// POUs/_FB_ConfigMachine
(****************************************************************************************************<br>
© Syntegon Group.<br>
All rights reserved, also regarding any disposal, exploitation, reproduction, editing, distribution,<br>
as well as in the event of applications for industrial property rights.<br>
*****************************************************************************************************<br>
DESCRIPTION:<br>
The machine as a whole (config protocol 3, ADR 0022): the recipe fields the application declares (process values<br>
such as belt speed, picks per cycle, the product pattern), their staging by the Simulator with the mechanism of the<br>
parameter sets, and the machine commands Start, Stop and Reset the application answers. One per application,<br>
listed in the config manifest with id 0. Typical cycle:<br>
  fb_Machine.m_Register(vio_Manifest := GVL_Config.stManifest, vi_udn_Id := 0);<br>
  fb_Machine.m_DeclareField(vi_un_Field := 1, vi_str_Name := 'BeltSpeed', vi_udn_Group := fb_Infeed.m_Id(),<br>
    vi_e_Type := E_ConfigFieldType.NUMBER, vi_str_Unit := 'mm/s', vi_lr_Min := 0, vi_lr_Max := 500,<br>
    vi_lr_ProgramValue := 150);<br>
  fb_Machine.m_SetText(vi_un_Field := 1, vi_str_Label := 'Belt speed', vi_str_Description := 'Speed of the infeed');<br>
  fb_Machine.m_SetVisibleWhen(vi_un_Field := 3, vi_un_OnField := 2, vi_dn_Value := 0);  // field 3 only with 2 = 0<br>
  fb_Machine.m_Cycle(vio_Set := RecipeSet, vi_b_ApplyAllowed := b_Stopped);<br>
  lr_BeltSpeed := fb_Machine.m_Value(vi_un_Field := 1);<br>
  CASE fb_Machine.m_Command() OF E_ConfigCommand.START: ...<br>
    fb_Machine.m_AnswerCommand(vi_b_Accepted := TRUE, vi_str_Reason := ''); END_CASE<br>
RecipeSet is the application's VAR PERSISTENT ST_ConfigRecipeSet.<br>
*****************************************************************************************************<br>
OUTPUT VALUES:<br>
vo_Config is the contract structure the gateway reads and writes at the path in the config manifest.<br>
*****************************************************************************************************<br>
LIMITS:<br>
CONFIG_un_MAX_RECIPE_FIELDS fields, CONFIG_un_MAX_CHOICES choices each. The gateway reads the declarations when<br>
it discovers the PLC: declare every field from the start and keep their order.<br>
*****************************************************************************************************<br>
VERSION         ¦ DATE       ¦ NAME      ¦ CHANGE<br>
Syn_Config 2.1.0 ¦ 2026-11-14 ¦ J.Willner ¦ Created: recipe fields and machine commands (protocol 3)<br>
Syn_Config 2.2.0 ¦ 2026-11-14 ¦ J.Willner ¦ m_SetText, m_SetVisibleWhen (protocol 4, #49)<br>
Syn_Config 2.3.0 ¦ 2026-11-14 ¦ J.Willner ¦ m_Cycle through m_HandleStaging<br>
****************************************************************************************************)
FUNCTION_BLOCK _FB_ConfigMachine EXTENDS _FB_ConfigComponent
VAR_OUTPUT
	vo_Config							: ST_ConfigMachine;	// contract structure of the gateway
END_VAR

(****************************************************************************************************<br>
© Syntegon Group.<br>
All rights reserved, also regarding any disposal, exploitation, reproduction, editing, distribution,<br>
as well as in the event of applications for industrial property rights.<br>
*****************************************************************************************************<br>
DESCRIPTION:<br>
Answers the waiting machine command: accepted, or rejected with the reason the Simulator shows. The command no<br>
longer waits afterwards.<br>
*****************************************************************************************************<br>
OUTPUT VALUES:<br>
FALSE while no command waits.<br>
****************************************************************************************************)
METHOD m_AnswerCommand : BOOL
VAR_INPUT
	vi_b_Accepted						: BOOL;	// TRUE: the application carries the command out
	vi_str_Reason						: STRING(80);	// why it is rejected, '' when accepted
END_VAR
m_AnswerCommand := vo_Config.stCommand.bRequested;
IF NOT m_AnswerCommand THEN
	RETURN;
END_IF
vo_Config.stCommandStatus.nHandledCommandId := vo_Config.stCommand.nCommandId;
vo_Config.stCommandStatus.eResult := SEL(vi_b_Accepted, E_ConfigCommandResult.REJECTED, E_ConfigCommandResult.ACCEPTED);
vo_Config.stCommandStatus.sMessage := SEL(vi_b_Accepted, vi_str_Reason, '');
vo_Config.stCommand.bRequested := FALSE;
END_METHOD

(****************************************************************************************************<br>
© Syntegon Group.<br>
All rights reserved, also regarding any disposal, exploitation, reproduction, editing, distribution,<br>
as well as in the event of applications for industrial property rights.<br>
*****************************************************************************************************<br>
DESCRIPTION:<br>
The machine command waiting for the application's answer (START, STOP, RESET); NONE while none waits. Answer it<br>
with m_AnswerCommand: the application alone decides whether it is carried out.<br>
****************************************************************************************************)
METHOD m_Command : E_ConfigCommand
IF vo_Config.stCommand.bRequested THEN
	m_Command := vo_Config.stCommand.eCommand;
ELSE
	m_Command := E_ConfigCommand.NONE;
END_IF
END_METHOD

(****************************************************************************************************<br>
© Syntegon Group.<br>
All rights reserved, also regarding any disposal, exploitation, reproduction, editing, distribution,<br>
as well as in the event of applications for industrial property rights.<br>
*****************************************************************************************************<br>
DESCRIPTION:<br>
Every cycle, after the fields are declared: handles a staged recipe or a reset (a recipe only while<br>
vi_b_ApplyAllowed), keeps the active recipe in vio_Set and gives the effective values in vo_Config.aActive: the<br>
active recipe while one is valid, else the fields' program values.<br>
*****************************************************************************************************<br>
OUTPUT VALUES:<br>
TRUE in the cycle a recipe was taken over or reset.<br>
****************************************************************************************************)
METHOD m_Cycle : BOOL
VAR_IN_OUT
	vio_Set								: ST_ConfigRecipeSet;	// the application's VAR PERSISTENT active recipe
END_VAR
VAR_INPUT
	vi_b_ApplyAllowed					: BOOL;	// [-] a staged recipe may be taken over now, e.g. while the machine stands
END_VAR
VAR
	b_TempTakeOver						: BOOL;	// the staged recipe was taken over: copy it
	un_TempIndex						: UINT;
END_VAR
m_Cycle := m_HandleStaging(vio_Staging := vo_Config.stStaging, vio_Status := vo_Config.stStatus, vio_b_Valid := vio_Set.bValid,
	vio_udn_Version := vio_Set.nVersion, vio_udn_LastVersion := vio_Set.nLastVersion, vi_b_ApplyAllowed := vi_b_ApplyAllowed,
	vo_b_TakeOver => b_TempTakeOver);
IF b_TempTakeOver THEN
	vio_Set.aValues := vo_Config.aStaged;
END_IF


(****************************************************************************************************
EFFECTIVE VALUES
****************************************************************************************************)
un_TempIndex := 0;
WHILE un_TempIndex < vo_Config.nFieldCount AND un_TempIndex < CONFIG_GlobalConst_Param.CONFIG_un_MAX_RECIPE_FIELDS DO
	vo_Config.aActive[un_TempIndex] := SEL(vio_Set.bValid, vo_Config.aFields[un_TempIndex].fProgramValue,
		vio_Set.aValues[un_TempIndex]);
	un_TempIndex := un_TempIndex + 1;
END_WHILE
END_METHOD

(****************************************************************************************************<br>
© Syntegon Group.<br>
All rights reserved, also regarding any disposal, exploitation, reproduction, editing, distribution,<br>
as well as in the event of applications for industrial property rights.<br>
*****************************************************************************************************<br>
DESCRIPTION:<br>
Declares recipe field vi_un_Field (1..CONFIG_un_MAX_RECIPE_FIELDS): its name, the component it belongs to, how its<br>
value is kept, its unit, range and the program value that applies while no recipe is active. Fields are listed up<br>
to the highest one declared. Idempotent: call it every cycle, before m_Cycle. A CHOICE field's values are named with<br>
m_SetChoice and range from 0; its vi_lr_Min and vi_lr_Max are not used, nor a SWITCH's.<br>
*****************************************************************************************************<br>
OUTPUT VALUES:<br>
FALSE for vi_un_Field = 0 or above CONFIG_un_MAX_RECIPE_FIELDS.<br>
****************************************************************************************************)
METHOD m_DeclareField : BOOL
VAR_INPUT
	vi_un_Field							: UINT;	// [-] 1..CONFIG_un_MAX_RECIPE_FIELDS
	vi_str_Name							: STRING(31);	// unique in the recipe, e.g. 'BeltSpeed'
	vi_udn_Group						: UDINT;	// [-] manifest id of the Syn_Visu component, 0 = the whole machine
	vi_e_Type							: E_ConfigFieldType;
	vi_str_Unit							: STRING(15);	// e.g. 'mm/s', '' = none
	vi_lr_Min							: LREAL;	// smallest value of a NUMBER or INTEGER field
	vi_lr_Max							: LREAL;	// largest value of a NUMBER or INTEGER field
	vi_lr_ProgramValue					: LREAL;	// the application's own value; a SWITCH: 1 = on
END_VAR
m_DeclareField := vi_un_Field > 0 AND vi_un_Field <= CONFIG_GlobalConst_Param.CONFIG_un_MAX_RECIPE_FIELDS;
IF NOT m_DeclareField THEN
	RETURN;
END_IF
vo_Config.aFields[vi_un_Field - 1].sName := vi_str_Name;
vo_Config.aFields[vi_un_Field - 1].nGroup := vi_udn_Group;
vo_Config.aFields[vi_un_Field - 1].eType := vi_e_Type;
vo_Config.aFields[vi_un_Field - 1].sUnit := vi_str_Unit;
vo_Config.aFields[vi_un_Field - 1].fMin := vi_lr_Min;
vo_Config.aFields[vi_un_Field - 1].fMax := vi_lr_Max;
vo_Config.aFields[vi_un_Field - 1].fProgramValue := vi_lr_ProgramValue;
IF vi_un_Field > vo_Config.nFieldCount THEN
	vo_Config.nFieldCount := vi_un_Field;
END_IF
END_METHOD

(****************************************************************************************************<br>
© Syntegon Group.<br>
All rights reserved, also regarding any disposal, exploitation, reproduction, editing, distribution,<br>
as well as in the event of applications for industrial property rights.<br>
*****************************************************************************************************<br>
DESCRIPTION:<br>
Effective value of an INTEGER or CHOICE recipe field as a whole number (see m_Value).<br>
****************************************************************************************************)
METHOD m_Integer : DINT
VAR_INPUT
	vi_un_Field							: UINT;	// [-] 1..the field count
END_VAR
m_Integer := LREAL_TO_DINT(m_Value(vi_un_Field := vi_un_Field));
END_METHOD

(****************************************************************************************************<br>
© Syntegon Group.<br>
All rights reserved, also regarding any disposal, exploitation, reproduction, editing, distribution,<br>
as well as in the event of applications for industrial property rights.<br>
*****************************************************************************************************<br>
DESCRIPTION:<br>
Why the staged recipe cannot be taken over; '' when it can: a value outside its field's range (NUMBER, INTEGER),<br>
not one of its choices (CHOICE), not a whole number (INTEGER, CHOICE) or not 0 or 1 (SWITCH).<br>
****************************************************************************************************)
METHOD PROTECTED m_InvalidStaged : STRING(80)
VAR
	un_TempIndex						: UINT;
	lr_TempValue						: LREAL;
	lr_TempMin							: LREAL;
	lr_TempMax							: LREAL;
END_VAR
m_InvalidStaged := '';
un_TempIndex := 0;
WHILE un_TempIndex < vo_Config.nFieldCount AND un_TempIndex < CONFIG_GlobalConst_Param.CONFIG_un_MAX_RECIPE_FIELDS DO
	lr_TempValue := vo_Config.aStaged[un_TempIndex];
	CASE vo_Config.aFields[un_TempIndex].eType OF
		E_ConfigFieldType.SWITCH:
			lr_TempMin := 0;
			lr_TempMax := 1;
		E_ConfigFieldType.CHOICE:
			lr_TempMin := 0;
			lr_TempMax := UINT_TO_LREAL(vo_Config.aFields[un_TempIndex].nChoiceCount) - 1;
	ELSE
		lr_TempMin := vo_Config.aFields[un_TempIndex].fMin;
		lr_TempMax := vo_Config.aFields[un_TempIndex].fMax;
	END_CASE
	(* The range first: only a value in range is turned into a whole number. NaN equals nothing, not even itself. *)
	IF lr_TempValue <> lr_TempValue OR lr_TempValue < lr_TempMin OR lr_TempValue > lr_TempMax THEN
		m_InvalidStaged := CONCAT(CONCAT('Field ', vo_Config.aFields[un_TempIndex].sName), CONCAT(': ', CONCAT(LREAL_TO_STRING(lr_TempValue),
			CONCAT(' is outside ', CONCAT(LREAL_TO_STRING(lr_TempMin), CONCAT(' to ', LREAL_TO_STRING(lr_TempMax)))))));
		RETURN;
	END_IF
	IF vo_Config.aFields[un_TempIndex].eType <> E_ConfigFieldType.NUMBER
		AND LINT_TO_LREAL(LREAL_TO_LINT(lr_TempValue)) <> lr_TempValue
	THEN
		m_InvalidStaged := CONCAT(CONCAT('Field ', vo_Config.aFields[un_TempIndex].sName), CONCAT(': ',
			CONCAT(LREAL_TO_STRING(lr_TempValue), ' is not a value of its type')));
		RETURN;
	END_IF
	un_TempIndex := un_TempIndex + 1;
END_WHILE
END_METHOD

(****************************************************************************************************<br>
© Syntegon Group.<br>
All rights reserved, also regarding any disposal, exploitation, reproduction, editing, distribution,<br>
as well as in the event of applications for industrial property rights.<br>
*****************************************************************************************************<br>
DESCRIPTION:<br>
Names value vi_un_Value (0..CONFIG_un_MAX_CHOICES-1) of the CHOICE field vi_un_Field, e.g. 0 = 'Lanes'. The field<br>
has as many choices as the highest value named plus one. Idempotent: call it every cycle with m_DeclareField.<br>
*****************************************************************************************************<br>
OUTPUT VALUES:<br>
FALSE for a field not declared or a value above CONFIG_un_MAX_CHOICES - 1.<br>
****************************************************************************************************)
METHOD m_SetChoice : BOOL
VAR_INPUT
	vi_un_Field							: UINT;	// [-] the field, 1..its count
	vi_un_Value							: UINT;	// [-] the value it names, from 0
	vi_str_Text							: STRING(31);	// e.g. 'Lanes'
END_VAR
m_SetChoice := vi_un_Field > 0 AND vi_un_Field <= vo_Config.nFieldCount
	AND vi_un_Value < CONFIG_GlobalConst_Param.CONFIG_un_MAX_CHOICES;
IF NOT m_SetChoice THEN
	RETURN;
END_IF
vo_Config.aFields[vi_un_Field - 1].aChoices[vi_un_Value] := vi_str_Text;
IF vi_un_Value >= vo_Config.aFields[vi_un_Field - 1].nChoiceCount THEN
	vo_Config.aFields[vi_un_Field - 1].nChoiceCount := vi_un_Value + 1;
END_IF
END_METHOD

(****************************************************************************************************<br>
© Syntegon Group.<br>
All rights reserved, also regarding any disposal, exploitation, reproduction, editing, distribution,<br>
as well as in the event of applications for industrial property rights.<br>
*****************************************************************************************************<br>
DESCRIPTION:<br>
Gives the declared field vi_un_Field the label the Simulator shows instead of its name put into words, and a<br>
description of what it is for, shown in the field's tooltip (config protocol 4, #49). Free text in the operators'<br>
language; the name stays the field's key. Idempotent: call it every cycle with m_DeclareField.<br>
*****************************************************************************************************<br>
OUTPUT VALUES:<br>
FALSE for a field not declared.<br>
****************************************************************************************************)
METHOD m_SetText : BOOL
VAR_INPUT
	vi_un_Field							: UINT;	// [-] the field, 1..its count
	vi_str_Label						: STRING(40);	// e.g. 'Belt speed', '' = the name put into words
	vi_str_Description					: STRING(160);	// what the field is for, '' = none
END_VAR
m_SetText := vi_un_Field > 0 AND vi_un_Field <= vo_Config.nFieldCount;
IF NOT m_SetText THEN
	RETURN;
END_IF
vo_Config.aFields[vi_un_Field - 1].sLabel := vi_str_Label;
vo_Config.aFields[vi_un_Field - 1].sDescription := vi_str_Description;
END_METHOD

(****************************************************************************************************<br>
© Syntegon Group.<br>
All rights reserved, also regarding any disposal, exploitation, reproduction, editing, distribution,<br>
as well as in the event of applications for industrial property rights.<br>
*****************************************************************************************************<br>
DESCRIPTION:<br>
Shows the declared field vi_un_Field in the Simulator only while field vi_un_OnField has the value vi_dn_Value<br>
(config protocol 4, #49), e.g. a lane count only while the pattern is Lanes. vi_un_OnField must be a SWITCH (0 / 1),<br>
CHOICE or INTEGER field and may belong to another group; a field depending on a hidden one is hidden too. A hidden<br>
field keeps its value and is written with the recipe. vi_un_OnField = 0 shows the field always. The gateway reports<br>
a condition on a NUMBER field, on the field itself, on a field not declared, on a value that field can never have<br>
or in a ring as a discovery error and shows that field always. Idempotent: call it every cycle with m_DeclareField.<br>
*****************************************************************************************************<br>
OUTPUT VALUES:<br>
FALSE for a field not declared.<br>
****************************************************************************************************)
METHOD m_SetVisibleWhen : BOOL
VAR_INPUT
	vi_un_Field							: UINT;	// [-] the field shown on condition, 1..its count
	vi_un_OnField						: UINT;	// [-] the field the condition reads, 0 = always shown
	vi_dn_Value							: DINT;	// [-] the value vi_un_OnField must have
END_VAR
m_SetVisibleWhen := vi_un_Field > 0 AND vi_un_Field <= vo_Config.nFieldCount;
IF NOT m_SetVisibleWhen THEN
	RETURN;
END_IF
vo_Config.aFields[vi_un_Field - 1].nVisibleField := vi_un_OnField;
vo_Config.aFields[vi_un_Field - 1].nVisibleValue := vi_dn_Value;
END_METHOD

(****************************************************************************************************<br>
© Syntegon Group.<br>
All rights reserved, also regarding any disposal, exploitation, reproduction, editing, distribution,<br>
as well as in the event of applications for industrial property rights.<br>
*****************************************************************************************************<br>
DESCRIPTION:<br>
Effective value of a SWITCH recipe field: TRUE for on (see m_Value).<br>
****************************************************************************************************)
METHOD m_Switch : BOOL
VAR_INPUT
	vi_un_Field							: UINT;	// [-] 1..the field count
END_VAR
m_Switch := m_Value(vi_un_Field := vi_un_Field) <> 0;
END_METHOD

(****************************************************************************************************<br>
© Syntegon Group.<br>
All rights reserved, also regarding any disposal, exploitation, reproduction, editing, distribution,<br>
as well as in the event of applications for industrial property rights.<br>
*****************************************************************************************************<br>
DESCRIPTION:<br>
Effective value of recipe field vi_un_Field, for the application's logic: the active recipe's, else the program<br>
value. 0 for a field not declared. A SWITCH gives 1 or 0, an INTEGER or CHOICE a whole number (m_Switch,<br>
m_Integer give them typed).<br>
****************************************************************************************************)
METHOD m_Value : LREAL
VAR_INPUT
	vi_un_Field							: UINT;	// [-] 1..the field count
END_VAR
IF vi_un_Field > 0 AND vi_un_Field <= vo_Config.nFieldCount THEN
	m_Value := vo_Config.aActive[vi_un_Field - 1];
ELSE
	m_Value := 0;
END_IF
END_METHOD

END_FUNCTION_BLOCK

// POUs/_FB_ConfigTopology
(****************************************************************************************************<br>
© Syntegon Group.<br>
All rights reserved, also regarding any disposal, exploitation, reproduction, editing, distribution,<br>
as well as in the event of applications for industrial property rights.<br>
*****************************************************************************************************<br>
DESCRIPTION:<br>
The machine's topology (config protocol 5, ADR 0023): how the parts of the application relate. The application<br>
declares the kinds of its topology nodes, the roles a link may have, every node of its full build-out with the<br>
Syn_Visu components it stands for, and its root node; its program values are the parents and links it uses. One per<br>
application, listed in the config manifest with id 0 like the machine FB. Typical cycle:<br>
  fb_Topology.m_Register(vio_Manifest := GVL_Config.stManifest, vi_udn_Id := 0);<br>
  fb_Topology.m_DeclareKind(vi_un_Kind := 1, vi_str_Name := 'Line');<br>
  fb_Topology.m_DeclareKind(vi_un_Kind := 2, vi_str_Name := 'PPH');<br>
  fb_Topology.m_AllowParent(vi_un_Kind := 2, vi_un_ParentKind := 1);<br>
  fb_Topology.m_DeclareRole(vi_un_Role := 1, vi_str_Name := 'Infeed1', vi_un_HolderKind := 2, vi_b_Required := TRUE);<br>
  fb_Topology.m_AllowTarget(vi_un_Role := 1, vi_un_TargetKind := 3);<br>
  fb_Topology.m_DeclareNode(vi_dn_Id := 21, vi_str_Name := 'PPH1', vi_un_Kind := 2);<br>
  fb_Topology.m_AddComponent(vi_dn_Node := 21, vi_udn_ComponentId := fb_Delta1.m_Id());<br>
  fb_Topology.m_SetRoot(vi_dn_Node := 1);<br>
  fb_Topology.m_SetParent(vi_dn_Node := 21, vi_dn_Parent := 1);<br>
  fb_Topology.m_Link(vi_dn_Node := 21, vi_un_Role := 1, vi_dn_Target := 30);<br>
  fb_Topology.m_Cycle();<br>
*****************************************************************************************************<br>
OUTPUT VALUES:<br>
vo_Config is the contract structure the gateway reads at the path in the config manifest.<br>
*****************************************************************************************************<br>
LIMITS:<br>
CONFIG_un_MAX_TOPOLOGY_KINDS kinds, CONFIG_un_MAX_TOPOLOGY_ROLES roles, CONFIG_un_MAX_TOPOLOGY_NODES nodes,<br>
CONFIG_un_MAX_TOPOLOGY_LINKS links, CONFIG_un_MAX_NODE_COMPONENTS components per node. The gateway reads the<br>
declaration when it discovers the PLC: declare everything from the start.<br>
*****************************************************************************************************<br>
VERSION         ¦ DATE       ¦ NAME      ¦ CHANGE<br>
Syn_Config 2.4.0 ¦ 2026-11-19 ¦ J.Willner ¦ Created: declaration and program values (protocol 5, #56)<br>
****************************************************************************************************)
FUNCTION_BLOCK _FB_ConfigTopology EXTENDS _FB_ConfigComponent
VAR_OUTPUT
	vo_Config							: ST_ConfigTopology;	// contract structure of the gateway
END_VAR
VAR
	ProgramLinks						: ST_ConfigTopologyLinks;	// the program values, given with m_SetParent and m_Link
END_VAR

(****************************************************************************************************<br>
© Syntegon Group.<br>
All rights reserved, also regarding any disposal, exploitation, reproduction, editing, distribution,<br>
as well as in the event of applications for industrial property rights.<br>
*****************************************************************************************************<br>
DESCRIPTION:<br>
Names a Syn_Visu component the declared node vi_dn_Node stands for, e.g. a PPH's Delta robot. Idempotent: call it<br>
every cycle with m_DeclareNode.<br>
*****************************************************************************************************<br>
OUTPUT VALUES:<br>
FALSE for a node not declared, component id 0, or more than CONFIG_un_MAX_NODE_COMPONENTS components.<br>
****************************************************************************************************)
METHOD m_AddComponent : BOOL
VAR_INPUT
	vi_dn_Node							: DINT;	// [-] the node's id
	vi_udn_ComponentId					: UDINT;	// [-] manifest id of the Syn_Visu component, e.g. fb_Delta1.m_Id()
END_VAR
VAR
	n_TempNode							: INT;
	un_TempIndex						: UINT;
END_VAR
n_TempNode := m_NodeIndex(vi_dn_Id := vi_dn_Node);
m_AddComponent := n_TempNode >= 0 AND vi_udn_ComponentId <> 0;
IF NOT m_AddComponent THEN
	RETURN;
END_IF
un_TempIndex := 0;
WHILE un_TempIndex < vo_Config.aNodes[n_TempNode].nComponentCount
	AND un_TempIndex < CONFIG_GlobalConst_Param.CONFIG_un_MAX_NODE_COMPONENTS
DO
	IF vo_Config.aNodes[n_TempNode].aComponents[un_TempIndex] = vi_udn_ComponentId THEN
		RETURN;
	END_IF
	un_TempIndex := un_TempIndex + 1;
END_WHILE
IF vo_Config.aNodes[n_TempNode].nComponentCount >= CONFIG_GlobalConst_Param.CONFIG_un_MAX_NODE_COMPONENTS THEN
	m_AddComponent := FALSE;
	RETURN;
END_IF
vo_Config.aNodes[n_TempNode].aComponents[vo_Config.aNodes[n_TempNode].nComponentCount] := vi_udn_ComponentId;
vo_Config.aNodes[n_TempNode].nComponentCount := vo_Config.aNodes[n_TempNode].nComponentCount + 1;
END_METHOD

(****************************************************************************************************<br>
© Syntegon Group.<br>
All rights reserved, also regarding any disposal, exploitation, reproduction, editing, distribution,<br>
as well as in the event of applications for industrial property rights.<br>
*****************************************************************************************************<br>
DESCRIPTION:<br>
Allows a node of kind vi_un_ParentKind to be the parent of a node of kind vi_un_Kind, e.g. a cell the parent of a<br>
PPH. Idempotent: call it every cycle with m_DeclareKind.<br>
*****************************************************************************************************<br>
OUTPUT VALUES:<br>
FALSE when either kind is not declared.<br>
****************************************************************************************************)
METHOD m_AllowParent : BOOL
VAR_INPUT
	vi_un_Kind							: UINT;	// [-] the child's kind, 1..its count
	vi_un_ParentKind					: UINT;	// [-] the parent's kind, 1..its count
END_VAR
m_AllowParent := vi_un_Kind > 0 AND vi_un_Kind <= vo_Config.nKindCount
	AND vi_un_ParentKind > 0 AND vi_un_ParentKind <= vo_Config.nKindCount;
IF NOT m_AllowParent THEN
	RETURN;
END_IF
vo_Config.aKinds[vi_un_Kind - 1].nParentKinds := vo_Config.aKinds[vi_un_Kind - 1].nParentKinds
	OR SHL(DWORD#1, vi_un_ParentKind - 1);
END_METHOD

(****************************************************************************************************<br>
© Syntegon Group.<br>
All rights reserved, also regarding any disposal, exploitation, reproduction, editing, distribution,<br>
as well as in the event of applications for industrial property rights.<br>
*****************************************************************************************************<br>
DESCRIPTION:<br>
Allows a link in role vi_un_Role to point to a node of kind vi_un_TargetKind, e.g. Infeed1 to a transport.<br>
Idempotent: call it every cycle with m_DeclareRole.<br>
*****************************************************************************************************<br>
OUTPUT VALUES:<br>
FALSE when the role or the kind is not declared.<br>
****************************************************************************************************)
METHOD m_AllowTarget : BOOL
VAR_INPUT
	vi_un_Role							: UINT;	// [-] the role, 1..its count
	vi_un_TargetKind					: UINT;	// [-] the kind it may point to, 1..its count
END_VAR
m_AllowTarget := vi_un_Role > 0 AND vi_un_Role <= vo_Config.nRoleCount
	AND vi_un_TargetKind > 0 AND vi_un_TargetKind <= vo_Config.nKindCount;
IF NOT m_AllowTarget THEN
	RETURN;
END_IF
vo_Config.aRoles[vi_un_Role - 1].nTargetKinds := vo_Config.aRoles[vi_un_Role - 1].nTargetKinds
	OR SHL(DWORD#1, vi_un_TargetKind - 1);
END_METHOD

(****************************************************************************************************<br>
© Syntegon Group.<br>
All rights reserved, also regarding any disposal, exploitation, reproduction, editing, distribution,<br>
as well as in the event of applications for industrial property rights.<br>
*****************************************************************************************************<br>
DESCRIPTION:<br>
Every cycle, after the declaration and the program values: gives the links in effect in vo_Config.stActive, the<br>
program values.<br>
*****************************************************************************************************<br>
OUTPUT VALUES:<br>
TRUE.<br>
****************************************************************************************************)
METHOD m_Cycle : BOOL
vo_Config.stActive := ProgramLinks;
m_Cycle := TRUE;
END_METHOD

(****************************************************************************************************<br>
© Syntegon Group.<br>
All rights reserved, also regarding any disposal, exploitation, reproduction, editing, distribution,<br>
as well as in the event of applications for industrial property rights.<br>
*****************************************************************************************************<br>
DESCRIPTION:<br>
Declares kind vi_un_Kind (1..CONFIG_un_MAX_TOPOLOGY_KINDS) of topology node, e.g. 'PPH' or 'Transport'. Kinds are<br>
listed up to the highest one declared. Idempotent: call it every cycle, before the roles and nodes.<br>
*****************************************************************************************************<br>
OUTPUT VALUES:<br>
FALSE for vi_un_Kind = 0 or above CONFIG_un_MAX_TOPOLOGY_KINDS.<br>
****************************************************************************************************)
METHOD m_DeclareKind : BOOL
VAR_INPUT
	vi_un_Kind							: UINT;	// [-] 1..CONFIG_un_MAX_TOPOLOGY_KINDS
	vi_str_Name							: STRING(31);	// unique in the topology, e.g. 'PPH'
END_VAR
m_DeclareKind := vi_un_Kind > 0 AND vi_un_Kind <= CONFIG_GlobalConst_Param.CONFIG_un_MAX_TOPOLOGY_KINDS;
IF NOT m_DeclareKind THEN
	RETURN;
END_IF
vo_Config.aKinds[vi_un_Kind - 1].sName := vi_str_Name;
IF vi_un_Kind > vo_Config.nKindCount THEN
	vo_Config.nKindCount := vi_un_Kind;
END_IF
END_METHOD

(****************************************************************************************************<br>
© Syntegon Group.<br>
All rights reserved, also regarding any disposal, exploitation, reproduction, editing, distribution,<br>
as well as in the event of applications for industrial property rights.<br>
*****************************************************************************************************<br>
DESCRIPTION:<br>
Declares the topology node vi_dn_Id of the full build-out, in use or not, with its name and kind; nodes are listed<br>
in the order they are first declared. Idempotent: call it every cycle, after m_DeclareKind.<br>
*****************************************************************************************************<br>
OUTPUT VALUES:<br>
FALSE for id 0, a kind not declared, or more than CONFIG_un_MAX_TOPOLOGY_NODES nodes.<br>
****************************************************************************************************)
METHOD m_DeclareNode : BOOL
VAR_INPUT
	vi_dn_Id							: DINT;	// [-] the application's id, e.g. its context id; not 0
	vi_str_Name							: STRING(31);	// e.g. 'PPH1'
	vi_un_Kind							: UINT;	// [-] its kind, 1..the kind count
END_VAR
VAR
	n_TempIndex							: INT;
END_VAR
m_DeclareNode := vi_dn_Id <> 0 AND vi_un_Kind > 0 AND vi_un_Kind <= vo_Config.nKindCount;
IF NOT m_DeclareNode THEN
	RETURN;
END_IF
n_TempIndex := m_NodeIndex(vi_dn_Id := vi_dn_Id);
IF n_TempIndex < 0 THEN
	IF vo_Config.nNodeCount >= CONFIG_GlobalConst_Param.CONFIG_un_MAX_TOPOLOGY_NODES THEN
		m_DeclareNode := FALSE;
		RETURN;
	END_IF
	n_TempIndex := UINT_TO_INT(vo_Config.nNodeCount);
	vo_Config.nNodeCount := vo_Config.nNodeCount + 1;
	vo_Config.aNodes[n_TempIndex].nId := vi_dn_Id;
END_IF
vo_Config.aNodes[n_TempIndex].sName := vi_str_Name;
vo_Config.aNodes[n_TempIndex].nKind := vi_un_Kind;
END_METHOD

(****************************************************************************************************<br>
© Syntegon Group.<br>
All rights reserved, also regarding any disposal, exploitation, reproduction, editing, distribution,<br>
as well as in the event of applications for industrial property rights.<br>
*****************************************************************************************************<br>
DESCRIPTION:<br>
Declares role vi_un_Role (1..CONFIG_un_MAX_TOPOLOGY_ROLES) a link may have, e.g. 'Infeed1' held by a PPH; the kinds<br>
it may point to are allowed with m_AllowTarget. Roles are listed up to the highest one declared. The parent is no<br>
role (m_SetParent). Idempotent: call it every cycle, after m_DeclareKind.<br>
*****************************************************************************************************<br>
OUTPUT VALUES:<br>
FALSE for vi_un_Role = 0 or above CONFIG_un_MAX_TOPOLOGY_ROLES, or a holder kind not declared.<br>
****************************************************************************************************)
METHOD m_DeclareRole : BOOL
VAR_INPUT
	vi_un_Role							: UINT;	// [-] 1..CONFIG_un_MAX_TOPOLOGY_ROLES
	vi_str_Name							: STRING(31);	// unique in the topology, e.g. 'Infeed1'
	vi_un_HolderKind					: UINT;	// [-] the kind of node that holds the role
	vi_b_Required						: BOOL;	// a node in use of that kind must have a link in this role
END_VAR
m_DeclareRole := vi_un_Role > 0 AND vi_un_Role <= CONFIG_GlobalConst_Param.CONFIG_un_MAX_TOPOLOGY_ROLES
	AND vi_un_HolderKind > 0 AND vi_un_HolderKind <= vo_Config.nKindCount;
IF NOT m_DeclareRole THEN
	RETURN;
END_IF
vo_Config.aRoles[vi_un_Role - 1].sName := vi_str_Name;
vo_Config.aRoles[vi_un_Role - 1].nHolderKind := vi_un_HolderKind;
vo_Config.aRoles[vi_un_Role - 1].bRequired := vi_b_Required;
IF vi_un_Role > vo_Config.nRoleCount THEN
	vo_Config.nRoleCount := vi_un_Role;
END_IF
END_METHOD

(****************************************************************************************************<br>
© Syntegon Group.<br>
All rights reserved, also regarding any disposal, exploitation, reproduction, editing, distribution,<br>
as well as in the event of applications for industrial property rights.<br>
*****************************************************************************************************<br>
DESCRIPTION:<br>
The topology is not staged yet (config protocol 5 has no topology staging): nothing to reject.<br>
****************************************************************************************************)
METHOD PROTECTED m_InvalidStaged : STRING(80)
m_InvalidStaged := '';
END_METHOD

(****************************************************************************************************<br>
© Syntegon Group.<br>
All rights reserved, also regarding any disposal, exploitation, reproduction, editing, distribution,<br>
as well as in the event of applications for industrial property rights.<br>
*****************************************************************************************************<br>
DESCRIPTION:<br>
A program value: node vi_dn_Node points to node vi_dn_Target in role vi_un_Role, e.g. PPH1's Infeed1 is TBL1. A<br>
node has one link per role; linking it again in that role replaces the target. Role 0 is the parent<br>
(m_SetParent). Idempotent: call it every cycle after the declaration, before m_Cycle.<br>
*****************************************************************************************************<br>
OUTPUT VALUES:<br>
FALSE for a node, target or role not declared, or more than CONFIG_un_MAX_TOPOLOGY_LINKS links.<br>
****************************************************************************************************)
METHOD m_Link : BOOL
VAR_INPUT
	vi_dn_Node							: DINT;	// [-] id of the node that holds the link
	vi_un_Role							: UINT;	// [-] its role, 1..the role count; 0 = the parent
	vi_dn_Target						: DINT;	// [-] id of the node it points to
END_VAR
VAR
	un_TempIndex						: UINT;
END_VAR
m_Link := m_NodeIndex(vi_dn_Id := vi_dn_Node) >= 0 AND m_NodeIndex(vi_dn_Id := vi_dn_Target) >= 0
	AND vi_un_Role <= vo_Config.nRoleCount;
IF NOT m_Link THEN
	RETURN;
END_IF

(* The node's link in this role, if it has one. *)
un_TempIndex := 0;
WHILE un_TempIndex < ProgramLinks.nLinkCount AND un_TempIndex < CONFIG_GlobalConst_Param.CONFIG_un_MAX_TOPOLOGY_LINKS DO
	IF ProgramLinks.aLinks[un_TempIndex].nNode = vi_dn_Node AND ProgramLinks.aLinks[un_TempIndex].nRole = vi_un_Role THEN
		ProgramLinks.aLinks[un_TempIndex].nTarget := vi_dn_Target;
		RETURN;
	END_IF
	un_TempIndex := un_TempIndex + 1;
END_WHILE

(* New link. *)
IF ProgramLinks.nLinkCount >= CONFIG_GlobalConst_Param.CONFIG_un_MAX_TOPOLOGY_LINKS THEN
	m_Link := FALSE;
	RETURN;
END_IF
ProgramLinks.aLinks[ProgramLinks.nLinkCount].nNode := vi_dn_Node;
ProgramLinks.aLinks[ProgramLinks.nLinkCount].nRole := vi_un_Role;
ProgramLinks.aLinks[ProgramLinks.nLinkCount].nTarget := vi_dn_Target;
ProgramLinks.nLinkCount := ProgramLinks.nLinkCount + 1;
END_METHOD

(****************************************************************************************************<br>
© Syntegon Group.<br>
All rights reserved, also regarding any disposal, exploitation, reproduction, editing, distribution,<br>
as well as in the event of applications for industrial property rights.<br>
*****************************************************************************************************<br>
DESCRIPTION:<br>
Index in vo_Config.aNodes of the node with id vi_dn_Id; -1 when none is declared.<br>
****************************************************************************************************)
METHOD PRIVATE m_NodeIndex : INT
VAR_INPUT
	vi_dn_Id							: DINT;	// [-] the node's id
END_VAR
VAR
	un_TempIndex						: UINT;
END_VAR
m_NodeIndex := -1;
un_TempIndex := 0;
WHILE un_TempIndex < vo_Config.nNodeCount AND un_TempIndex < CONFIG_GlobalConst_Param.CONFIG_un_MAX_TOPOLOGY_NODES DO
	IF vo_Config.aNodes[un_TempIndex].nId = vi_dn_Id THEN
		m_NodeIndex := UINT_TO_INT(un_TempIndex);
		RETURN;
	END_IF
	un_TempIndex := un_TempIndex + 1;
END_WHILE
END_METHOD

(****************************************************************************************************<br>
© Syntegon Group.<br>
All rights reserved, also regarding any disposal, exploitation, reproduction, editing, distribution,<br>
as well as in the event of applications for industrial property rights.<br>
*****************************************************************************************************<br>
DESCRIPTION:<br>
A program value: node vi_dn_Parent is the parent of node vi_dn_Node (m_Link in role 0). Idempotent: call it every<br>
cycle after the declaration, before m_Cycle.<br>
*****************************************************************************************************<br>
OUTPUT VALUES:<br>
FALSE as m_Link.<br>
****************************************************************************************************)
METHOD m_SetParent : BOOL
VAR_INPUT
	vi_dn_Node							: DINT;	// [-] id of the child
	vi_dn_Parent						: DINT;	// [-] id of its parent
END_VAR
m_SetParent := m_Link(vi_dn_Node := vi_dn_Node, vi_un_Role := 0, vi_dn_Target := vi_dn_Parent);
END_METHOD

(****************************************************************************************************<br>
© Syntegon Group.<br>
All rights reserved, also regarding any disposal, exploitation, reproduction, editing, distribution,<br>
as well as in the event of applications for industrial property rights.<br>
*****************************************************************************************************<br>
DESCRIPTION:<br>
Makes the declared node vi_dn_Node the root node: the one node without a parent, from which every node in use<br>
hangs. Idempotent: call it every cycle after m_DeclareNode. A topology has one root node: another one is refused.<br>
*****************************************************************************************************<br>
OUTPUT VALUES:<br>
FALSE for a node not declared, or a second root node.<br>
****************************************************************************************************)
METHOD m_SetRoot : BOOL
VAR_INPUT
	vi_dn_Node							: DINT;	// [-] the node's id
END_VAR
m_SetRoot := m_NodeIndex(vi_dn_Id := vi_dn_Node) >= 0
	AND (vo_Config.nRootNode = 0 OR vo_Config.nRootNode = vi_dn_Node);
IF m_SetRoot THEN
	vo_Config.nRootNode := vi_dn_Node;
END_IF
END_METHOD

END_FUNCTION_BLOCK

// POUs/_FB_ConfigCartesian
(****************************************************************************************************<br>
© Syntegon Group.<br>
All rights reserved, also regarding any disposal, exploitation, reproduction, editing, distribution,<br>
as well as in the event of applications for industrial property rights.<br>
*****************************************************************************************************<br>
DESCRIPTION:<br>
Parameter set of one Cartesian robot (ADR 0017): its pose, origin shift, zones, gripper fingers, limit area and<br>
TCP limit area, written by the configurator, taken over when the application allows it.<br>
Typical cycle:<br>
  fb_CartParam.m_Register(vio_Manifest := GVL_Config.stManifest, vi_udn_Id := fb_Cart.m_Id());<br>
  fb_CartParam.m_Cycle(vio_Default := CartDefault, vio_Set := CartSet, vi_b_ApplyAllowed := b_Stopped);<br>
  fb_Cart.m_Configure(vi_lr_XMin := 0, ...);<br>
  fb_CartParam.m_PassOn(vio_Visu := fb_Cart);<br>
The application's logic takes its zones and limit areas from m_Active, not from its own constants.<br>
*****************************************************************************************************<br>
OUTPUT VALUES:<br>
vo_Config is the contract structure the gateway reads and writes at the path in the config manifest.<br>
*****************************************************************************************************<br>
VERSION         ¦ DATE       ¦ NAME      ¦ CHANGE<br>
Syn_Config 1.1.0 ¦ 2026-11-10 ¦ J.Willner ¦ New<br>
Syn_Config 2.0.0 ¦ 2026-11-11 ¦ J.Willner ¦ Gripper fingers with their offsets, m_Invalid (ADR 0018)<br>
Syn_Config 2.3.0 ¦ 2026-11-14 ¦ J.Willner ¦ m_Cycle through m_HandleStaging; m_PassOn passes the pose on<br>
****************************************************************************************************)
FUNCTION_BLOCK _FB_ConfigCartesian EXTENDS _FB_ConfigComponent
VAR_OUTPUT
	vo_Config							: ST_ConfigCartesian;	// contract structure of the gateway
END_VAR

(****************************************************************************************************<br>
© Syntegon Group.<br>
All rights reserved, also regarding any disposal, exploitation, reproduction, editing, distribution,<br>
as well as in the event of applications for industrial property rights.<br>
*****************************************************************************************************<br>
DESCRIPTION:<br>
All effective values (zones, limit areas, ...), for the application's own logic.<br>
****************************************************************************************************)
METHOD m_Active : ST_ConfigCartesianParam
m_Active := vo_Config.stActive;
END_METHOD

(****************************************************************************************************<br>
© Syntegon Group.<br>
All rights reserved, also regarding any disposal, exploitation, reproduction, editing, distribution,<br>
as well as in the event of applications for industrial property rights.<br>
*****************************************************************************************************<br>
DESCRIPTION:<br>
A Cartesian robot.<br>
****************************************************************************************************)
METHOD PROTECTED m_ComponentType : SynVisu.E_VisuComponentType
m_ComponentType := SynVisu.E_VisuComponentType.CARTESIAN;
END_METHOD

(****************************************************************************************************<br>
© Syntegon Group.<br>
All rights reserved, also regarding any disposal, exploitation, reproduction, editing, distribution,<br>
as well as in the event of applications for industrial property rights.<br>
*****************************************************************************************************<br>
DESCRIPTION:<br>
Every cycle: handles a staged set or a reset (a set only while vi_b_ApplyAllowed), keeps the active set in<br>
vio_Set and gives the effective values in vo_Config.stActive: the active set while one is valid, else the<br>
program values vio_Default.<br>
*****************************************************************************************************<br>
OUTPUT VALUES:<br>
TRUE in the cycle a set was taken over or reset.<br>
****************************************************************************************************)
METHOD m_Cycle : BOOL
VAR_IN_OUT CONSTANT
	vio_Default							: ST_ConfigCartesianParam;	// the application's program values
END_VAR
VAR_IN_OUT
	vio_Set								: ST_ConfigCartesianSet;	// the application's VAR PERSISTENT active set
END_VAR
VAR_INPUT
	vi_b_ApplyAllowed					: BOOL;	// [-] a staged set may be taken over now, e.g. while the machine stands
END_VAR
VAR
	b_TempTakeOver						: BOOL;	// the staged set was taken over: copy it
END_VAR
m_Cycle := m_HandleStaging(vio_Staging := vo_Config.stStaging, vio_Status := vo_Config.stStatus, vio_b_Valid := vio_Set.bValid,
	vio_udn_Version := vio_Set.nVersion, vio_udn_LastVersion := vio_Set.nLastVersion, vi_b_ApplyAllowed := vi_b_ApplyAllowed,
	vo_b_TakeOver => b_TempTakeOver);
IF b_TempTakeOver THEN
	vio_Set.stParam := vo_Config.stStaged;
END_IF


(****************************************************************************************************
EFFECTIVE VALUES
****************************************************************************************************)
IF vio_Set.bValid THEN
	vo_Config.stActive := vio_Set.stParam;
ELSE
	vo_Config.stActive := vio_Default;
END_IF
END_METHOD

(****************************************************************************************************<br>
© Syntegon Group.<br>
All rights reserved, also regarding any disposal, exploitation, reproduction, editing, distribution,<br>
as well as in the event of applications for industrial property rights.<br>
*****************************************************************************************************<br>
DESCRIPTION:<br>
Why a staged set cannot be taken over; '' when it can: more zones or fingers than the lists hold, a zone on no<br>
conveyor (id 0), or a finger without a diameter or height.<br>
****************************************************************************************************)
METHOD PROTECTED m_InvalidStaged : STRING(80)
m_InvalidStaged := m_InvalidZones(vio_aZones := vo_Config.stStaged.aZones, vi_un_Count := vo_Config.stStaged.nZoneCount);
IF m_InvalidStaged = '' THEN
	m_InvalidStaged := m_InvalidFingers(vio_aFingers := vo_Config.stStaged.aFingers, vi_un_Count := vo_Config.stStaged.nFingerCount);
END_IF
END_METHOD

(****************************************************************************************************<br>
© Syntegon Group.<br>
All rights reserved, also regarding any disposal, exploitation, reproduction, editing, distribution,<br>
as well as in the event of applications for industrial property rights.<br>
*****************************************************************************************************<br>
DESCRIPTION:<br>
Passes the effective pose, origin shift, limit areas, zones and fingers on to the robot's Syn_Visu FB, so the<br>
visualisation shows what the machine uses; the strokes and rail height (hardware) stay with the application's<br>
m_Configure call. Call it after m_Cycle, every cycle; Syn_Visu's config version only changes when a value does.<br>
****************************************************************************************************)
METHOD m_PassOn : BOOL
VAR_IN_OUT
	vio_Visu							: SynVisu._FB_VisuCartesian;	// the robot's Syn_Visu FB
END_VAR
m_PassOn := TRUE;
vio_Visu.m_SetPose(vi_Pose := vo_Config.stActive.stPose);
vio_Visu.m_SetOriginShift(vi_lr_X := vo_Config.stActive.stOriginShift.fX, vi_lr_Y := vo_Config.stActive.stOriginShift.fY,
	vi_lr_Z := vo_Config.stActive.stOriginShift.fZ);
m_PassOnLimitAreas(vio_Visu := vio_Visu, vio_LimitArea := vo_Config.stActive.stLimitArea,
	vio_TcpLimitArea := vo_Config.stActive.stTcpLimitArea);
m_PassOnZones(vio_Visu := vio_Visu, vio_aZones := vo_Config.stActive.aZones, vi_un_Count := vo_Config.stActive.nZoneCount,
	vi_un_VisuCount := vio_Visu.vo_Visu.stConfig.nZoneCount);
m_PassOnFingers(vio_Visu := vio_Visu, vio_aFingers := vo_Config.stActive.aFingers,
	vi_un_Count := vo_Config.stActive.nFingerCount, vi_un_VisuCount := vio_Visu.vo_Visu.stConfig.nFingerCount);
END_METHOD

(****************************************************************************************************<br>
© Syntegon Group.<br>
All rights reserved, also regarding any disposal, exploitation, reproduction, editing, distribution,<br>
as well as in the event of applications for industrial property rights.<br>
*****************************************************************************************************<br>
DESCRIPTION:<br>
Effective pose of the axis origin (MCS), for the application's logic.<br>
****************************************************************************************************)
METHOD m_Pose : SynVisu.ST_VisuPose
m_Pose := vo_Config.stActive.stPose;
END_METHOD

END_FUNCTION_BLOCK

// POUs/_FB_ConfigXtsLoop
(****************************************************************************************************<br>
© Syntegon Group.<br>
All rights reserved, also regarding any disposal, exploitation, reproduction, editing, distribution,<br>
as well as in the event of applications for industrial property rights.<br>
*****************************************************************************************************<br>
DESCRIPTION:<br>
Parameter set of one XTS loop (ADR 0017): its pose, origin shift, track modules, zones and gripper fingers,<br>
written by the configurator, taken over when the application allows it. Typical cycle:<br>
  fb_FxxParam.m_Register(vio_Manifest := GVL_Config.stManifest, vi_udn_Id := fb_Fxx.m_Id());<br>
  fb_FxxParam.m_Cycle(vio_Default := FxxDefault, vio_Set := FxxSet, vi_b_ApplyAllowed := b_Stopped);<br>
  fb_Fxx.m_Configure(vi_lr_ToolOffset := 120, ...);<br>
  fb_FxxParam.m_PassOn(vio_Visu := fb_Fxx);<br>
The application's logic takes its track and zones from m_Active, not from its own constants.<br>
*****************************************************************************************************<br>
OUTPUT VALUES:<br>
vo_Config is the contract structure the gateway reads and writes at the path in the config manifest.<br>
*****************************************************************************************************<br>
VERSION         ¦ DATE       ¦ NAME      ¦ CHANGE<br>
Syn_Config 1.1.0 ¦ 2026-11-10 ¦ J.Willner ¦ New<br>
Syn_Config 2.0.0 ¦ 2026-11-11 ¦ J.Willner ¦ Gripper fingers with their offsets (ADR 0018)<br>
Syn_Config 2.3.0 ¦ 2026-11-14 ¦ J.Willner ¦ m_Cycle through m_HandleStaging; m_PassOn passes the pose on<br>
****************************************************************************************************)
FUNCTION_BLOCK _FB_ConfigXtsLoop EXTENDS _FB_ConfigComponent
VAR_OUTPUT
	vo_Config							: ST_ConfigXtsLoop;	// contract structure of the gateway
END_VAR

(****************************************************************************************************<br>
© Syntegon Group.<br>
All rights reserved, also regarding any disposal, exploitation, reproduction, editing, distribution,<br>
as well as in the event of applications for industrial property rights.<br>
*****************************************************************************************************<br>
DESCRIPTION:<br>
All effective values (track modules, zones, ...), for the application's own logic.<br>
****************************************************************************************************)
METHOD m_Active : ST_ConfigXtsLoopParam
m_Active := vo_Config.stActive;
END_METHOD

(****************************************************************************************************<br>
© Syntegon Group.<br>
All rights reserved, also regarding any disposal, exploitation, reproduction, editing, distribution,<br>
as well as in the event of applications for industrial property rights.<br>
*****************************************************************************************************<br>
DESCRIPTION:<br>
An XTS loop.<br>
****************************************************************************************************)
METHOD PROTECTED m_ComponentType : SynVisu.E_VisuComponentType
m_ComponentType := SynVisu.E_VisuComponentType.XTS_LOOP;
END_METHOD

(****************************************************************************************************<br>
© Syntegon Group.<br>
All rights reserved, also regarding any disposal, exploitation, reproduction, editing, distribution,<br>
as well as in the event of applications for industrial property rights.<br>
*****************************************************************************************************<br>
DESCRIPTION:<br>
Every cycle: handles a staged set or a reset (a set only while vi_b_ApplyAllowed), keeps the active set in<br>
vio_Set and gives the effective values in vo_Config.stActive: the active set while one is valid, else the<br>
program values vio_Default.<br>
*****************************************************************************************************<br>
OUTPUT VALUES:<br>
TRUE in the cycle a set was taken over or reset.<br>
****************************************************************************************************)
METHOD m_Cycle : BOOL
VAR_IN_OUT CONSTANT
	vio_Default							: ST_ConfigXtsLoopParam;	// the application's program values
END_VAR
VAR_IN_OUT
	vio_Set								: ST_ConfigXtsLoopSet;	// the application's VAR PERSISTENT active set
END_VAR
VAR_INPUT
	vi_b_ApplyAllowed					: BOOL;	// [-] a staged set may be taken over now, e.g. while the machine stands
END_VAR
VAR
	b_TempTakeOver						: BOOL;	// the staged set was taken over: copy it
END_VAR
m_Cycle := m_HandleStaging(vio_Staging := vo_Config.stStaging, vio_Status := vo_Config.stStatus, vio_b_Valid := vio_Set.bValid,
	vio_udn_Version := vio_Set.nVersion, vio_udn_LastVersion := vio_Set.nLastVersion, vi_b_ApplyAllowed := vi_b_ApplyAllowed,
	vo_b_TakeOver => b_TempTakeOver);
IF b_TempTakeOver THEN
	vio_Set.stParam := vo_Config.stStaged;
END_IF


(****************************************************************************************************
EFFECTIVE VALUES
****************************************************************************************************)
IF vio_Set.bValid THEN
	vo_Config.stActive := vio_Set.stParam;
ELSE
	vo_Config.stActive := vio_Default;
END_IF
END_METHOD

(****************************************************************************************************<br>
© Syntegon Group.<br>
All rights reserved, also regarding any disposal, exploitation, reproduction, editing, distribution,<br>
as well as in the event of applications for industrial property rights.<br>
*****************************************************************************************************<br>
DESCRIPTION:<br>
Why a staged set cannot be taken over; '' when it can: a track without modules, more modules, zones or fingers<br>
than the lists hold, a module without a length, a zone on no conveyor (id 0), or a finger without a diameter or<br>
height.<br>
****************************************************************************************************)
METHOD PROTECTED m_InvalidStaged : STRING(80)
m_InvalidStaged := m_InvalidModules(vio_aModules := vo_Config.stStaged.aModules, vi_un_Count := vo_Config.stStaged.nModuleCount);
IF m_InvalidStaged = '' THEN
	m_InvalidStaged := m_InvalidZones(vio_aZones := vo_Config.stStaged.aZones, vi_un_Count := vo_Config.stStaged.nZoneCount);
END_IF
IF m_InvalidStaged = '' THEN
	m_InvalidStaged := m_InvalidFingers(vio_aFingers := vo_Config.stStaged.aFingers, vi_un_Count := vo_Config.stStaged.nFingerCount);
END_IF
END_METHOD

(****************************************************************************************************<br>
© Syntegon Group.<br>
All rights reserved, also regarding any disposal, exploitation, reproduction, editing, distribution,<br>
as well as in the event of applications for industrial property rights.<br>
*****************************************************************************************************<br>
DESCRIPTION:<br>
Passes the effective pose, origin shift, track modules, zones and fingers on to the loop's Syn_Visu FB, so the<br>
visualisation shows what the machine uses; the tool offset and mover size (hardware) stay with the<br>
application's m_Configure call. Call it after m_Cycle, every cycle; Syn_Visu's config version only changes when<br>
a value does.<br>
****************************************************************************************************)
METHOD m_PassOn : BOOL
VAR_IN_OUT
	vio_Visu							: SynVisu._FB_VisuXtsLoop;	// the loop's Syn_Visu FB
END_VAR
m_PassOn := TRUE;
vio_Visu.m_SetPose(vi_Pose := vo_Config.stActive.stPose);
vio_Visu.m_SetOriginShift(vi_lr_X := vo_Config.stActive.stOriginShift.fX, vi_lr_Y := vo_Config.stActive.stOriginShift.fY,
	vi_lr_Z := vo_Config.stActive.stOriginShift.fZ);
m_PassOnModules(vio_Visu := vio_Visu, vio_aModules := vo_Config.stActive.aModules,
	vi_un_Count := vo_Config.stActive.nModuleCount, vi_un_VisuCount := vio_Visu.vo_Visu.stConfig.nModuleCount);
m_PassOnZones(vio_Visu := vio_Visu, vio_aZones := vo_Config.stActive.aZones, vi_un_Count := vo_Config.stActive.nZoneCount,
	vi_un_VisuCount := vio_Visu.vo_Visu.stConfig.nZoneCount);
m_PassOnFingers(vio_Visu := vio_Visu, vio_aFingers := vo_Config.stActive.aFingers,
	vi_un_Count := vo_Config.stActive.nFingerCount, vi_un_VisuCount := vio_Visu.vo_Visu.stConfig.nFingerCount);
END_METHOD

(****************************************************************************************************<br>
© Syntegon Group.<br>
All rights reserved, also regarding any disposal, exploitation, reproduction, editing, distribution,<br>
as well as in the event of applications for industrial property rights.<br>
*****************************************************************************************************<br>
DESCRIPTION:<br>
Effective pose of the start of module 1 (MCS), for the application's logic.<br>
****************************************************************************************************)
METHOD m_Pose : SynVisu.ST_VisuPose
m_Pose := vo_Config.stActive.stPose;
END_METHOD

END_FUNCTION_BLOCK

// POUs/_FC_GetVersionSynConfig
(****************************************************************************************************<br>
© Syntegon Group.<br>
All rights reserved, also regarding any disposal, exploitation, reproduction, editing, distribution,<br>
as well as in the event of applications for industrial property rights.<br>
*****************************************************************************************************<br>
DESCRIPTION:<br>
Runtime-readable version of the Syn_Config library.<br>
*****************************************************************************************************<br>
VERSION         ¦ DATE       ¦ NAME      ¦ CHANGE<br>
Syn_Config 1.0.0 ¦ 2026-11-10 ¦ J.Willner ¦ Parameter sets of conveyors and Deltas (ADR 0017, protocol 1)<br>
Syn_Config 1.1.0 ¦ 2026-11-10 ¦ J.Willner ¦ Every other component type (#24)<br>
Syn_Config 2.0.0 ¦ 2026-11-11 ¦ J.Willner ¦ Gripper fingers in the robots' sets (protocol 2, #25)<br>
Syn_Config 2.0.1 ¦ 2026-11-12 ¦ J.Willner ¦ SynVisu as a placeholder: the application chooses its version<br>
Syn_Config 2.1.0 ¦ 2026-11-14 ¦ J.Willner ¦ Machine FB: recipe fields and machine commands (protocol 3, #43)<br>
Syn_Config 2.2.0 ¦ 2026-11-14 ¦ J.Willner ¦ Recipe fields: label, description, visibility condition (protocol 4, #49)<br>
Syn_Config 2.3.0 ¦ 2026-11-14 ¦ J.Willner ¦ One staging lifecycle; m_PassOn passes the pose on (Syn_Visu 10.0.0)<br>
Syn_Config 2.4.0 ¦ 2026-11-19 ¦ J.Willner ¦ Topology FB: nodes, roles and program links (protocol 5, #56)<br>
****************************************************************************************************)
FUNCTION _FC_GetVersionSynConfig : UINT
VAR_INPUT
	vi_n_VersionElement					: INT;	// [-] 1 = major, 2 = minor, 3 = revision
END_VAR

CASE vi_n_VersionElement OF
	1: _FC_GetVersionSynConfig := 2;
	2: _FC_GetVersionSynConfig := 4;
	3: _FC_GetVersionSynConfig := 0;
ELSE
	_FC_GetVersionSynConfig := 16#FFFF;
END_CASE

END_FUNCTION
